{attribute 'qualified_only'}
{attribute 'strict'}
{attribute 'to_string'}
TYPE E_MBDataType :
(
    mbNone      := 0,
    mbReal32    := 1,
    mbInt32     := 2,
    mbUInt32    := 3,
    mbInt16     := 4,
    mbUInt16    := 5,
    mbWord16    := 6,
    mbBit       := 7
) UINT;
END_TYPE

(* stored: Version 1.1.0.1
   DUT E_MBDataType: Id {610641d5-177b-4292-a8fe-cea258ced114} *)
